// TIA Portal V21 export
// export: Created 2026-11-10T19:21:31.8595839Z, ExportSetting WithDefaults, DisplayName Totally Integrated Automation Portal, DisplayVersion V21 Update 3, DisplayName STEP 7 Professional, DisplayVersion V21 Update 3, DisplayName STEP 7 Safety, DisplayVersion V21, DisplayName Tech WebApplication, DisplayVersion V21, DisplayName WinCC Basic/Comfort/Advanced, DisplayVersion V21 Update 3, DisplayName WinCC Unified, DisplayVersion V21 Update 3
FUNCTION_BLOCK "FB_Lad_mb002"   // FB7, LAD
{ S7_Optimized_Access := 'TRUE' }
VERSION : 0.1
// stored: AutoNumber true, IsIECCheckEnabled false, IsRetainMemResEnabled false, MemoryReserve 100, SetENOAutomatically false, UDAEnableTagReadback false
   VAR_INPUT
      v_req : Bool;
      v_mb_addr : UInt;
      v_mode : USInt;
      v_data_addr : UDInt;
      v_data_len : UInt;
   END_VAR
   VAR_OUTPUT
      v_done : Bool;
      v_busy : Bool;
      v_error : Bool;
      v_status : Word;
   END_VAR
   VAR_IN_OUT
      v_data_ptr : Variant;
   END_VAR
   VAR
      inst { S7_SetPoint := 'True'} : Modbus_Master;
   END_VAR
BEGIN

REGION Network 1: Description of MB_MASTER
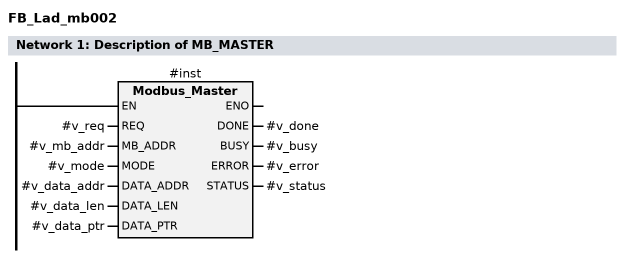
   RUNG wire#powerrail
      #inst.Modbus_Master(REQ := #v_req, MB_ADDR := #v_mb_addr, MODE := #v_mode, DATA_ADDR := #v_data_addr, DATA_LEN := #v_data_len, DONE => #v_done, BUSY => #v_busy, ERROR => #v_error, STATUS => #v_status, DATA_PTR := #v_data_ptr)
   END_RUNG
   // the same network as SCL:
   #inst(REQ := #v_req,   // Modbus_Master
         MB_ADDR := #v_mb_addr,
         MODE := #v_mode,
         DATA_ADDR := #v_data_addr,
         DATA_LEN := #v_data_len,
         DATA_PTR := #v_data_ptr,
         DONE => #v_done,
         BUSY => #v_busy,
         ERROR => #v_error,
         STATUS => #v_status);
END_REGION
END_FUNCTION_BLOCK
